(* IEC 61131-3 sources: Versio-VersionControlSystem/fixtures/projects/RefrigeratorControl/Device/Plc Logic/Application/Library/Alarm/DUTs/Hmi, 1 file *)

(* ---- ST_AlarmHmiConfiguration.st ---- *)
//{attribute 'OPC' := '2'}
TYPE ST_AlarmHmiConfiguration :
STRUCT
	Info			: STRING(40); // PL use instead
	Initialized		: BOOL;
END_STRUCT
END_TYPE
